RoboDK station: simulation.rdk

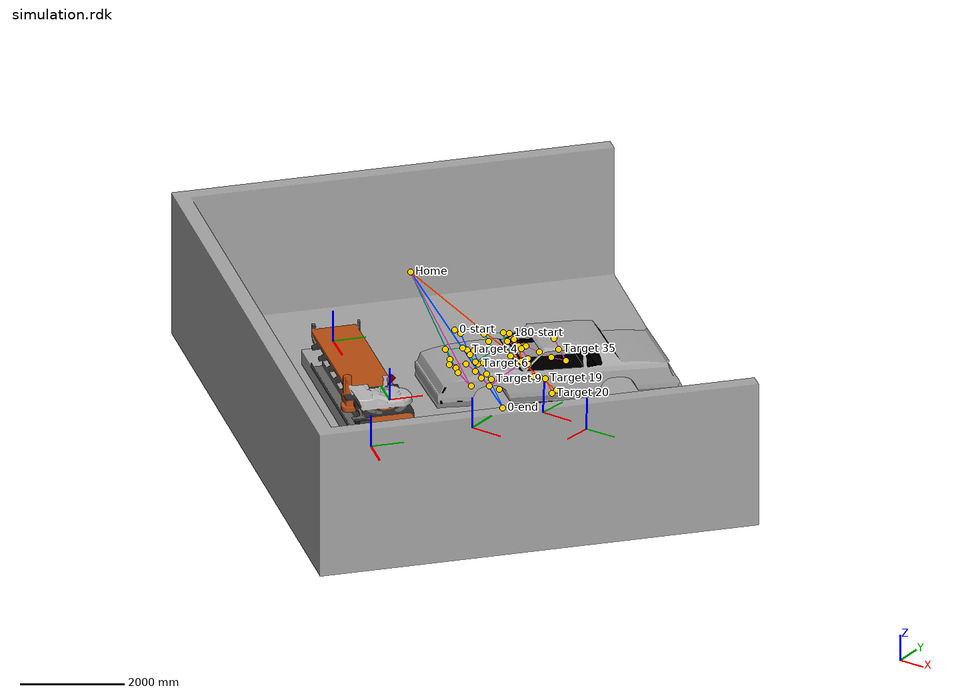
[picture v0: the station drawn from its stored meshes, robots at their saved joint values, targets as dots, program paths as lines]
Station New Station (1)2 (saved by RoboDK 6.1.1). Poses are relative to the parent item; angles as X-Y-Z fixed-axis rotations.
  - frame Frame 1 at (0, 0, 0) mm
    - frame Turn Table Base at (1090.8, 803.58, 313.71) mm, rotated rx -3.83 ry -0.12 rz 0.01 deg
      - robot Turn Table: 1 axes
          modified DH rows (alpha deg, a mm, theta deg, d mm): 0, 0, 0, 0
          joint limits [-360] to [360]; home [0]; saved at [270]
        - frame Frame 5 at (-0.07, 1018.58, -71.28) mm, rotated rx 0.95 ry 0 rz 0.22 deg
        - tool internship 2, TCP at (0, 0, 200) mm, size 4802.1 x 1035.2 x 1720.5 mm, geometry from internship 2.STL
      - target turn_0 (joint target) at (0, 0, 200) mm; joints [0] of Turn Table
      - target turn_90 (joint target) at (0, 0, 200) mm, rotated rx 0 ry 0 rz 90 deg; joints [90] of Turn Table
      - target turn_180 (joint target) at (0, 0, 200) mm, rotated rx 0 ry 0 rz 180 deg; joints [180] of Turn Table
      - target turn_270 (joint target) at (0, 0, 200) mm, rotated rx 0 ry 0 rz -90 deg; joints [270] of Turn Table
    - object layout2 at (0, 0, 0) mm, rotated rx 90 ry 0 rz 140 deg, size 11000 x 3000 x 8700 mm, geometry from layout2.STL
  - frame Frame 6 at (0, -3390, 970) mm, rotated rx 0 ry 0 rz -40 deg
    - object base at (-1330, 140, 0) mm, rotated rx 90 ry 0 rz 0 deg, size 5000 x 300 x 1000 mm, geometry from base.STL
  - frame ABB IRBT 6004 Standard 3.5m Base at (-2780, -680, 1350) mm, rotated rx 0 ry 0 rz -39.7 deg
    - robot ABB IRBT 6004 Standard 3.5m: 1 axes, repeatability 0.1 mm
        modified DH rows (alpha deg, a mm, theta deg, d mm): 0, 0, 0, 0 linear
        base shift (840.5, 4.2, 379.5) mm, rotated rx 0 ry 90 rz 0 deg
        joint limits [0] to [3500]; home [0]; saved at [2827.078]
      - frame ABB IRB 6650S-90/3.9 Base at (-160, 160, 0) mm, rotated rx -2.54 ry 0.52 rz 90 deg
        - robot ABB IRB 6650S-90/3.9: 6 axes, payload 90 kg, reach 3900 mm, repeatability 0.14 mm, weight 2275 kg
            joint limits [-180, -40, -180, -300, -120, -360] to [180, 160, 70, 300, 120, 360]; home [0, 0, 0, 0, 0, 0]; saved at [-94.567, -9.168, -174.099, 70.725, 70.561, 76.601]
          - tool Paint gun, TCP at (50, -150, 740) mm, rotated rx 0 ry 30 rz 0 deg, size 203.2 x 279.7 x 471.5 mm
        - target Home (joint target) at (926.35, 1847.38, 1781.69) mm, rotated rx -116.33 ry 65.1 rz -108.86 deg; joints [-94.567, -9.168, -174.099, 70.725, 70.561, 76.601] of ABB IRB 6650S-90/3.9
        - target 0-start (Cartesian target) at (2184.4, 3279.5, -176.12) mm, rotated rx -96.51 ry 63.32 rz -79.51 deg; joints [65.271, 78.343, -26.977, 31.951, -81.109, -50.329] of ABB IRB 6650S-90/3.9
        - target Target 3 (Cartesian target) at (2165.69, 2792.62, -41.51) mm, rotated rx -96.51 ry 63.32 rz -79.51 deg; joints [61.504, 60.223, 1.958, 28.188, -89.439, -43.105] of ABB IRB 6650S-90/3.9
        - target Target 4 (Cartesian target) at (2155.28, 2226.68, -153.05) mm, rotated rx -96.51 ry 63.32 rz -79.51 deg; joints [55.139, 54.811, 20.629, 22.886, -100.409, -35.301] of ABB IRB 6650S-90/3.9
        - target Target 5 (Cartesian target) at (2191.78, 1902.7, -29.79) mm, rotated rx -96.51 ry 63.32 rz -79.51 deg; joints [49.311, 45.605, 32.857, 17.675, -102.785, -32.974] of ABB IRB 6650S-90/3.9
        - target Target 6 (Cartesian target) at (2168.89, 1506.86, -146.21) mm, rotated rx -96.51 ry 63.32 rz -79.51 deg; joints [41.711, 48.218, 39.943, 11.122, -111.941, -29.557] of ABB IRB 6650S-90/3.9
        - target Target 7 (Cartesian target) at (2186.24, 1201.33, 6.36) mm, rotated rx -96.51 ry 63.32 rz -79.51 deg; joints [33.345, 38.15, 50.265, 2.874, -112.162, -29.257] of ABB IRB 6650S-90/3.9
        - target Target 8 (Cartesian target) at (2142.01, 813.18, -61.09) mm, rotated rx -96.51 ry 63.32 rz -79.51 deg; joints [21.226, 41.741, 54.511, -9.733, -119.912, -30.322] of ABB IRB 6650S-90/3.9
        - target Target 9 (Cartesian target) at (2127.2, 390.29, 9.13) mm, rotated rx -96.51 ry 63.32 rz -79.51 deg; joints [4.097, 36.802, 60.091, -27.932, -119.881, -32.691] of ABB IRB 6650S-90/3.9
        - target Target 10 (Cartesian target) at (2165.79, -57.5, -12.41) mm, rotated rx -96.51 ry 63.32 rz -79.51 deg; joints [-14.615, 38.345, 57.062, -46.92, -117.504, -33.482] of ABB IRB 6650S-90/3.9
        - target 0-end (Cartesian target) at (2112.66, -486.82, -218.44) mm, rotated rx -96.51 ry 63.32 rz -79.51 deg; joints [-31.008, 51.535, 46.37, -64.821, -117.323, -36.985] of ABB IRB 6650S-90/3.9
        - target 180-start (Cartesian target) at (3190.24, 2993.58, -241.99) mm, rotated rx -134.64 ry 54.92 rz -136.14 deg; joints [53.739, 102.57, -78.062, 65.937, -54.325, -80.517] of ABB IRB 6650S-90/3.9
        - target Target 13 (Cartesian target) at (3197.13, 2670.72, -227.94) mm, rotated rx -134.64 ry 54.92 rz -136.14 deg; joints [50.557, 79.011, -38.527, 54.328, -59.998, -62.423] of ABB IRB 6650S-90/3.9
        - target Target 14 (Cartesian target) at (3188.72, 2314.84, -214.93) mm, rotated rx -134.64 ry 54.92 rz -136.14 deg; joints [46.702, 67.154, -18.013, 47.05, -63.371, -52.846] of ABB IRB 6650S-90/3.9
        - target Target 15 (Cartesian target) at (3101.58, 1800.08, -311.55) mm, rotated rx -134.64 ry 54.92 rz -136.14 deg; joints [40.864, 58.009, 3.108, 37.674, -69.98, -41.383] of ABB IRB 6650S-90/3.9
        - target Target 16 (Cartesian target) at (3101.38, 1307.16, -172.22) mm, rotated rx -134.64 ry 54.92 rz -136.14 deg; joints [32.467, 45.569, 19.642, 28.276, -71.345, -35.659] of ABB IRB 6650S-90/3.9
        - target Target 17 (Cartesian target) at (3102.52, 896.64, -258.24) mm, rotated rx -134.64 ry 54.92 rz -136.14 deg; joints [24.005, 44.954, 26.053, 18.857, -75.387, -30.23] of ABB IRB 6650S-90/3.9
        - target Target 18 (Cartesian target) at (3117.33, 510.53, -115.48) mm, rotated rx -134.64 ry 54.92 rz -136.14 deg; joints [14.804, 36.206, 33.765, 9.426, -73.635, -27.403] of ABB IRB 6650S-90/3.9
        - target Target 19 (Cartesian target) at (3125.83, 147.97, 6.43) mm, rotated rx -134.64 ry 54.92 rz -136.14 deg; joints [5.526, 29.243, 38.382, -0.233, -71.034, -24.093] of ABB IRB 6650S-90/3.9
        - target Target 20 (Cartesian target) at (3125.54, -354.26, -84.61) mm, rotated rx -134.64 ry 54.92 rz -136.14 deg; joints [-7.629, 33.735, 36.285, -13.901, -73.981, -19.465] of ABB IRB 6650S-90/3.9
        - target 180-end (Cartesian target) at (3124.63, -677.04, 108.76) mm, rotated rx -134.64 ry 54.92 rz -136.14 deg; joints [-15.765, 26.511, 36.997, -23.112, -68.834, -14.079] of ABB IRB 6650S-90/3.9
        - target 270-start (Cartesian target) at (2840.07, 1218.88, -115.24) mm, rotated rx -169.44 ry 8.59 rz -153.99 deg; joints [29.407, 14.901, 28.49, 125.206, -13.821, -128.636] of ABB IRB 6650S-90/3.9
        - target Target 23 (Cartesian target) at (2883.32, 1763.75, -162) mm, rotated rx -169.44 ry 8.59 rz -153.99 deg; joints [38.43, 28.895, 12.077, 125.204, -20.683, -122.294] of ABB IRB 6650S-90/3.9
        - target Target 24 (Cartesian target) at (2883.7, 2301.08, 95.96) mm, rotated rx -169.44 ry 8.59 rz -153.99 deg; joints [45.86, 37.294, -7.912, 138.562, -32.981, -132.374] of ABB IRB 6650S-90/3.9
        - target Target 25 (Cartesian target) at (2576.82, 2561.47, 2.09) mm, rotated rx -169.44 ry 8.59 rz -153.99 deg; joints [52.955, 39.028, -7.493, 133.517, -35.689, -121.915] of ABB IRB 6650S-90/3.9
        - target Target 26 (Cartesian target) at (2539.75, 2081.36, 43.52) mm, rotated rx -169.44 ry 8.59 rz -153.99 deg; joints [47.742, 22.554, 13.621, 129.679, -29.372, -120.814] of ABB IRB 6650S-90/3.9
        - target Target 27 (Cartesian target) at (2463, 1571.27, 55.47) mm, rotated rx -169.44 ry 8.59 rz -153.99 deg; joints [41.019, 5.744, 33.047, 128.242, -23.58, -123.781] of ABB IRB 6650S-90/3.9
        - target Target 28 (Cartesian target) at (2085.21, 1417.27, -52.32) mm, rotated rx -169.44 ry 8.59 rz -153.99 deg; joints [44.681, -8.232, 50.464, 120.583, -23.934, -112.817] of ABB IRB 6650S-90/3.9
        - target Target 29 (Cartesian target) at (2098.76, 1871.89, -96.26) mm, rotated rx -169.44 ry 8.59 rz -153.99 deg; joints [52.152, 8.914, 34.782, 117.59, -28.012, -103.828] of ABB IRB 6650S-90/3.9
        - target Target 30 (Cartesian target) at (2089.73, 2335.43, -146.04) mm, rotated rx -169.44 ry 8.59 rz -153.99 deg; joints [58.153, 24.695, 17.184, 120.713, -32.742, -102.721] of ABB IRB 6650S-90/3.9
        - target Target 31 (Cartesian target) at (1803.93, 2561.24, -231.74) mm, rotated rx -169.44 ry 8.59 rz -153.99 deg; joints [65.441, 29.364, 13.854, 120.057, -36.702, -95.929] of ABB IRB 6650S-90/3.9
        - target Target 32 (Cartesian target) at (1732.63, 1975.31, -186.88) mm, rotated rx -169.44 ry 8.59 rz -153.99 deg; joints [60.98, 7.291, 39.887, 113.814, -32.105, -92.205] of ABB IRB 6650S-90/3.9
        - target 270-end (Cartesian target) at (1703.95, 1425.37, -136.41) mm, rotated rx -169.44 ry 8.59 rz -153.99 deg; joints [53.342, -18.383, 61.735, 118.225, -28.936, -103.618] of ABB IRB 6650S-90/3.9
        - target 90-start (Cartesian target) at (3684.29, 1522.85, 201.99) mm, rotated rx -177.66 ry 18.93 rz -162.21 deg; joints [26.55, 40.441, -13.305, 148.757, -16.778, -145.215] of ABB IRB 6650S-90/3.9
        - target Target 35 (Cartesian target) at (3659.36, 1089.59, 165.94) mm, rotated rx -177.66 ry 18.93 rz -162.21 deg; joints [19.677, 32.958, -1.68, 160.564, -10.413, -160.79] of ABB IRB 6650S-90/3.9
        - target Target 36 (Cartesian target) at (3651.01, 569.4, 142.24) mm, rotated rx -177.66 ry 18.93 rz -162.21 deg; joints [10.341, 27.714, 6.161, 206.471, -8.08, -212.307] of ABB IRB 6650S-90/3.9
        - target Target 37 (Cartesian target) at (3356.15, 525.98, 267.26) mm, rotated rx -177.66 ry 18.93 rz -162.21 deg; joints [10.558, 13.148, 20.355, 204.358, -8.338, -210.05] of ABB IRB 6650S-90/3.9
        - target Target 38 (Cartesian target) at (3233.88, 980.27, 202.02) mm, rotated rx -177.66 ry 18.93 rz -162.21 deg; joints [20.53, 14.764, 20.54, 144.903, -7.128, -144.477] of ABB IRB 6650S-90/3.9
        - target Target 39 (Cartesian target) at (3101.99, 1463.95, 137.32) mm, rotated rx -177.66 ry 18.93 rz -162.21 deg; joints [30.803, 19.872, 16.427, 115.861, -13.113, -108.941] of ABB IRB 6650S-90/3.9
        - target Target 40 (Cartesian target) at (2748.04, 1484.65, 271.41) mm, rotated rx -177.66 ry 18.93 rz -162.21 deg; joints [35.345, 5.095, 29.18, 118.828, -17.334, -109.297] of ABB IRB 6650S-90/3.9
        - target Target 41 (Cartesian target) at (2888.39, 1005.95, 308.2) mm, rotated rx -177.66 ry 18.93 rz -162.21 deg; joints [24.002, -0.85, 34.116, 140.167, -10.496, -137.709] of ABB IRB 6650S-90/3.9
        - target Target 42 (Cartesian target) at (2893.16, 538.55, 290.33) mm, rotated rx -177.66 ry 18.93 rz -162.21 deg; joints [13.029, -7.15, 40.67, 191.801, -7.678, -195.994] of ABB IRB 6650S-90/3.9
        - target Target 43 (Cartesian target) at (2057.36, 313.62, -95.92) mm, rotated rx -177.32 ry -4.8 rz -163.72 deg; joints [13.373, -34.598, 66.696, -1.997, 32.613, -2.29] of ABB IRB 6650S-90/3.9
        - target Target 44 (Cartesian target) at (2041.84, 816.3, -129.35) mm, rotated rx -177.32 ry -4.8 rz -163.72 deg; joints [28.595, -21.19, 58.837, -15.597, 28.992, 23.601] of ABB IRB 6650S-90/3.9
        - target Target 45 (Cartesian target) at (2029.36, 1228.07, -156.75) mm, rotated rx -177.32 ry -4.8 rz -163.72 deg; joints [38.698, -7.905, 48.971, -24.767, 28.481, 41.347] of ABB IRB 6650S-90/3.9
        - target Target 46 (Cartesian target) at (1966.11, 1668.4, -182.69) mm, rotated rx -177.32 ry -4.8 rz -163.72 deg; joints [48.074, 4.745, 37.486, -30.438, 30.711, 55.025] of ABB IRB 6650S-90/3.9
        - target Target 47 (Cartesian target) at (1633.89, 1663.16, -159.92) mm, rotated rx -177.32 ry -4.8 rz -163.72 deg; joints [54.611, -5.557, 46.943, -31.975, 33.962, 62] of ABB IRB 6650S-90/3.9
        - target Target 48 (Cartesian target) at (1680.61, 1169.79, -129.23) mm, rotated rx -177.32 ry -4.8 rz -163.72 deg; joints [44.216, -26.672, 62.693, -24.3, 34.862, 44.839] of ABB IRB 6650S-90/3.9
        - target 90-end (Cartesian target) at (1846.1, 837.14, -287.79) mm, rotated rx -177.32 ry -4.8 rz -163.72 deg; joints [32.332, -24.633, 66.62, -21.113, 25.769, 32.503] of ABB IRB 6650S-90/3.9
  - program 0 (11 instructions, listed below)
  - program 180 (13 instructions, listed below)
  - program 270 (15 instructions, listed below)
  - program 90 (19 instructions, listed below)
  - program main (10 instructions, listed below)
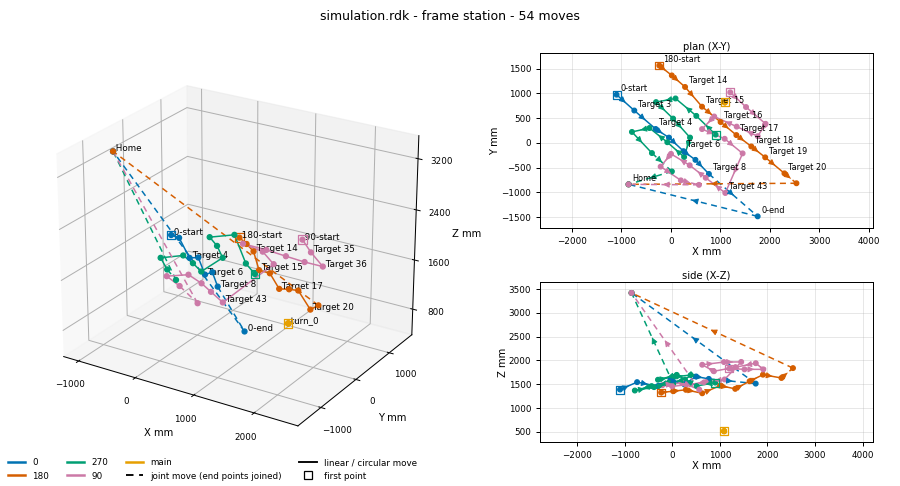
[picture p0: tool path of simulation.rdk in frame station, 54 of 54 moves have a stored position in this frame; points joined in program order, loops and branches not executed]

--- program 0 (robot ABB IRB 6650S-90/3.9) ---
  Set Ref.: ABB IRB 6650S-90/3.9 Base
  Set Tool: Paint gun
  MoveJ (0-start)
  MoveL (Target 3)
  MoveL (Target 4)
  MoveL (Target 5)
  MoveL (Target 6)
  MoveL (Target 7)
  MoveL (Target 8)
  MoveJ (0-end)
  MoveJ (Home)

--- program 180 (robot ABB IRB 6650S-90/3.9) ---
  Set Ref.: ABB IRB 6650S-90/3.9 Base
  Set Tool: Paint gun
  MoveJ (180-start)
  MoveL (Target 13)
  MoveL (Target 14)
  MoveL (Target 15)
  MoveL (Target 16)
  MoveL (Target 17)
  MoveL (Target 18)
  MoveL (Target 19)
  MoveL (Target 20)
  MoveJ (180-end)
  MoveJ (Home)

--- program 270 (robot ABB IRB 6650S-90/3.9) ---
  Set Ref.: ABB IRB 6650S-90/3.9 Base
  Set Tool: Paint gun
  MoveJ (270-start)
  MoveL (Target 23)
  MoveL (Target 24)
  MoveL (Target 25)
  MoveL (Target 26)
  MoveL (Target 27)
  MoveL (Target 28)
  MoveL (Target 29)
  MoveL (Target 30)
  MoveL (Target 31)
  MoveL (Target 32)
  MoveJ (270-end)
  MoveJ (Home)

--- program 90 (robot ABB IRB 6650S-90/3.9) ---
  Set Ref.: ABB IRB 6650S-90/3.9 Base
  Set Tool: Paint gun
  MoveJ (90-start)
  MoveL (Target 35)
  MoveL (Target 36)
  MoveL (Target 37)
  MoveL (Target 38)
  MoveL (Target 39)
  MoveL (Target 40)
  MoveL (Target 41)
  MoveL (Target 42)
  MoveL (Target 43)
  MoveL (Target 44)
  MoveL (Target 45)
  MoveL (Target 46)
  MoveL (Target 47)
  MoveL (Target 48)
  MoveJ (90-end)
  MoveJ (Home)

--- program main (robot Turn Table) ---
  Set Ref.: Turn Table Base
  Set Tool: internship 2
  MoveJ (turn_0)
  Call 0
  MoveJ (turn_90)
  Call 90
  MoveJ (turn_180)
  Call 180
  MoveJ (turn_270)
  Call 270
